(* IEC 61131-3 sources: s7-to-codesys/tests/POUs/Scenarios/FB_AnalogIn_ScenarioTest, 7 files *)

(* ---- FB_AnalogIn_ScenarioTest.decl.st ---- *)
// AUTO-GENERATED — не редактировать: s7conv gen-tests, сценарии scenarios/FB_AnalogIn.csv
// Правка — в CSV (scenarios/README.md), затем python -m s7conv build-corpus.
// Назначение: тесты поведения сконвертированного FB_AnalogIn по сценариям CSV (сценариев: 6, строк: 47):
//             один метод-тест на сценарий, строки — по порядку с моделируемым временем GVL_S7Clock.
//             Ожидаемые значения — из CSV (эталонные модели по описанию логики блока), не из
//             результата конвертации.
// Автор:      s7conv 0.1.0 (сгенерировано)
// Версия:     не указана
// Документ:   scenarios/README.md, docs/methodology.md, раздел «Проверка поведения»
FUNCTION_BLOCK FB_AnalogIn_ScenarioTest EXTENDS coUnit.FB_TestSuite
VAR
    fbScalingPoints : FB_AnalogIn;  // свой экземпляр на сценарий
    xScalingPointsDone : BOOL;  // сценарий выполнен (выполняется один раз)
    fbHighLimitsHysteresis : FB_AnalogIn;  // свой экземпляр на сценарий
    xHighLimitsHysteresisDone : BOOL;  // сценарий выполнен (выполняется один раз)
    fbLowLimitsHysteresis : FB_AnalogIn;  // свой экземпляр на сценарий
    xLowLimitsHysteresisDone : BOOL;  // сценарий выполнен (выполняется один раз)
    fbChannelDiagnostics : FB_AnalogIn;  // свой экземпляр на сценарий
    xChannelDiagnosticsDone : BOOL;  // сценарий выполнен (выполняется один раз)
    fbSimulation : FB_AnalogIn;  // свой экземпляр на сценарий
    xSimulationDone : BOOL;  // сценарий выполнен (выполняется один раз)
    fbCustomRanges : FB_AnalogIn;  // свой экземпляр на сценарий
    xCustomRangesDone : BOOL;  // сценарий выполнен (выполняется один раз)
END_VAR

(* ---- ChannelDiagnostics.method.impl.st ---- *)
// AUTO-GENERATED — не редактировать: scenarios/FB_AnalogIn.csv, сценарий ChannelDiagnostics
coUnit.TEST('ChannelDiagnostics');
IF NOT xChannelDiagnosticsDone THEN
    xChannelDiagnosticsDone := TRUE;
    GVL_S7Clock.xSimulation := TRUE;

    // #1, t = 0 мс — норма 8.0; замещающее значение 5.0
    GVL_S7Clock.tSimNow := T#0MS;
    fbChannelDiagnostics.raw := 13824;
    fbChannelDiagnostics.rangeLow := 0.0;
    fbChannelDiagnostics.rangeHigh := 16.0;
    fbChannelDiagnostics.limitHH := 14.0;
    fbChannelDiagnostics.limitH := 12.0;
    fbChannelDiagnostics.limitL := 2.0;
    fbChannelDiagnostics.limitLL := 1.0;
    fbChannelDiagnostics.hysteresis := 0.5;
    fbChannelDiagnostics.substitute := 5.0;
    fbChannelDiagnostics.simulation := FALSE;
    fbChannelDiagnostics.simValue := 0.0;
    fbChannelDiagnostics();
    AssertEquals_REAL(Expected := 8.0,
                      Actual := fbChannelDiagnostics.value,
                      Delta := 0.001,
                      Message := 'ChannelDiagnostics#1 value');
    AssertEquals_BOOL(Expected := TRUE, Actual := fbChannelDiagnostics.valid, Message := 'ChannelDiagnostics#1 valid');
    AssertEquals_BOOL(Expected := FALSE,
                      Actual := fbChannelDiagnostics.channelFault,
                      Message := 'ChannelDiagnostics#1 channelFault');
    AssertEquals_BOOL(Expected := FALSE,
                      Actual := fbChannelDiagnostics.overrange,
                      Message := 'ChannelDiagnostics#1 overrange');
    AssertEquals_BOOL(Expected := FALSE,
                      Actual := fbChannelDiagnostics.underrange,
                      Message := 'ChannelDiagnostics#1 underrange');
    AssertEquals_BOOL(Expected := FALSE,
                      Actual := fbChannelDiagnostics.alarmHH,
                      Message := 'ChannelDiagnostics#1 alarmHH');
    AssertEquals_BOOL(Expected := FALSE, Actual := fbChannelDiagnostics.warnH, Message := 'ChannelDiagnostics#1 warnH');
    AssertEquals_BOOL(Expected := FALSE, Actual := fbChannelDiagnostics.warnL, Message := 'ChannelDiagnostics#1 warnL');
    AssertEquals_BOOL(Expected := FALSE,
                      Actual := fbChannelDiagnostics.alarmLL,
                      Message := 'ChannelDiagnostics#1 alarmLL');
    AssertEquals_WORD(Expected := 16#0001,
                      Actual := fbChannelDiagnostics.statusWord,
                      Message := 'ChannelDiagnostics#1 statusWord');

    // #2, t = 100 мс — выше номинала: overrange, value ограничено 16.0, HH и H
    GVL_S7Clock.tSimNow := T#100MS;
    fbChannelDiagnostics.raw := 27649;
    fbChannelDiagnostics();
    AssertEquals_REAL(Expected := 16.0,
                      Actual := fbChannelDiagnostics.value,
                      Delta := 0.001,
                      Message := 'ChannelDiagnostics#2 value');
    AssertEquals_BOOL(Expected := TRUE, Actual := fbChannelDiagnostics.valid, Message := 'ChannelDiagnostics#2 valid');
    AssertEquals_BOOL(Expected := FALSE,
                      Actual := fbChannelDiagnostics.channelFault,
                      Message := 'ChannelDiagnostics#2 channelFault');
    AssertEquals_BOOL(Expected := TRUE,
                      Actual := fbChannelDiagnostics.overrange,
                      Message := 'ChannelDiagnostics#2 overrange');
    AssertEquals_BOOL(Expected := FALSE,
                      Actual := fbChannelDiagnostics.underrange,
                      Message := 'ChannelDiagnostics#2 underrange');
    AssertEquals_BOOL(Expected := TRUE,
                      Actual := fbChannelDiagnostics.alarmHH,
                      Message := 'ChannelDiagnostics#2 alarmHH');
    AssertEquals_BOOL(Expected := TRUE, Actual := fbChannelDiagnostics.warnH, Message := 'ChannelDiagnostics#2 warnH');
    AssertEquals_BOOL(Expected := FALSE, Actual := fbChannelDiagnostics.warnL, Message := 'ChannelDiagnostics#2 warnL');
    AssertEquals_BOOL(Expected := FALSE,
                      Actual := fbChannelDiagnostics.alarmLL,
                      Message := 'ChannelDiagnostics#2 alarmLL');
    AssertEquals_WORD(Expected := 16#0035,
                      Actual := fbChannelDiagnostics.statusWord,
                      Message := 'ChannelDiagnostics#2 statusWord');

    // #3, t = 200 мс — верхняя граница зоны перегрузки — ещё не неисправность
    GVL_S7Clock.tSimNow := T#200MS;
    fbChannelDiagnostics.raw := 32511;
    fbChannelDiagnostics();
    AssertEquals_REAL(Expected := 16.0,
                      Actual := fbChannelDiagnostics.value,
                      Delta := 0.001,
                      Message := 'ChannelDiagnostics#3 value');
    AssertEquals_BOOL(Expected := TRUE, Actual := fbChannelDiagnostics.valid, Message := 'ChannelDiagnostics#3 valid');
    AssertEquals_BOOL(Expected := FALSE,
                      Actual := fbChannelDiagnostics.channelFault,
                      Message := 'ChannelDiagnostics#3 channelFault');
    AssertEquals_BOOL(Expected := TRUE,
                      Actual := fbChannelDiagnostics.overrange,
                      Message := 'ChannelDiagnostics#3 overrange');
    AssertEquals_BOOL(Expected := FALSE,
                      Actual := fbChannelDiagnostics.underrange,
                      Message := 'ChannelDiagnostics#3 underrange');
    AssertEquals_BOOL(Expected := TRUE,
                      Actual := fbChannelDiagnostics.alarmHH,
                      Message := 'ChannelDiagnostics#3 alarmHH');
    AssertEquals_BOOL(Expected := TRUE, Actual := fbChannelDiagnostics.warnH, Message := 'ChannelDiagnostics#3 warnH');
    AssertEquals_BOOL(Expected := FALSE, Actual := fbChannelDiagnostics.warnL, Message := 'ChannelDiagnostics#3 warnL');
    AssertEquals_BOOL(Expected := FALSE,
                      Actual := fbChannelDiagnostics.alarmLL,
                      Message := 'ChannelDiagnostics#3 alarmLL');
    AssertEquals_WORD(Expected := 16#0035,
                      Actual := fbChannelDiagnostics.statusWord,
                      Message := 'ChannelDiagnostics#3 statusWord');

    // #4, t = 300 мс — за зоной перегрузки: channelFault, value := substitute, уставки сброшены
    GVL_S7Clock.tSimNow := T#300MS;
    fbChannelDiagnostics.raw := 32512;
    fbChannelDiagnostics();
    AssertEquals_REAL(Expected := 5.0,
                      Actual := fbChannelDiagnostics.value,
                      Delta := 0.001,
                      Message := 'ChannelDiagnostics#4 value');
    AssertEquals_BOOL(Expected := FALSE, Actual := fbChannelDiagnostics.valid, Message := 'ChannelDiagnostics#4 valid');
    AssertEquals_BOOL(Expected := TRUE,
                      Actual := fbChannelDiagnostics.channelFault,
                      Message := 'ChannelDiagnostics#4 channelFault');
    AssertEquals_BOOL(Expected := FALSE,
                      Actual := fbChannelDiagnostics.overrange,
                      Message := 'ChannelDiagnostics#4 overrange');
    AssertEquals_BOOL(Expected := FALSE,
                      Actual := fbChannelDiagnostics.underrange,
                      Message := 'ChannelDiagnostics#4 underrange');
    AssertEquals_BOOL(Expected := FALSE,
                      Actual := fbChannelDiagnostics.alarmHH,
                      Message := 'ChannelDiagnostics#4 alarmHH');
    AssertEquals_BOOL(Expected := FALSE, Actual := fbChannelDiagnostics.warnH, Message := 'ChannelDiagnostics#4 warnH');
    AssertEquals_BOOL(Expected := FALSE, Actual := fbChannelDiagnostics.warnL, Message := 'ChannelDiagnostics#4 warnL');
    AssertEquals_BOOL(Expected := FALSE,
                      Actual := fbChannelDiagnostics.alarmLL,
                      Message := 'ChannelDiagnostics#4 alarmLL');
    AssertEquals_WORD(Expected := 16#0002,
                      Actual := fbChannelDiagnostics.statusWord,
                      Message := 'ChannelDiagnostics#4 statusWord');

    // #5, t = 400 мс — переполнение/обрыв (7FFF)
    GVL_S7Clock.tSimNow := T#400MS;
    fbChannelDiagnostics.raw := 32767;
    fbChannelDiagnostics();
    AssertEquals_REAL(Expected := 5.0,
                      Actual := fbChannelDiagnostics.value,
                      Delta := 0.001,
                      Message := 'ChannelDiagnostics#5 value');
    AssertEquals_BOOL(Expected := FALSE, Actual := fbChannelDiagnostics.valid, Message := 'ChannelDiagnostics#5 valid');
    AssertEquals_BOOL(Expected := TRUE,
                      Actual := fbChannelDiagnostics.channelFault,
                      Message := 'ChannelDiagnostics#5 channelFault');
    AssertEquals_BOOL(Expected := FALSE,
                      Actual := fbChannelDiagnostics.overrange,
                      Message := 'ChannelDiagnostics#5 overrange');
    AssertEquals_BOOL(Expected := FALSE,
                      Actual := fbChannelDiagnostics.underrange,
                      Message := 'ChannelDiagnostics#5 underrange');
    AssertEquals_BOOL(Expected := FALSE,
                      Actual := fbChannelDiagnostics.alarmHH,
                      Message := 'ChannelDiagnostics#5 alarmHH');
    AssertEquals_BOOL(Expected := FALSE, Actual := fbChannelDiagnostics.warnH, Message := 'ChannelDiagnostics#5 warnH');
    AssertEquals_BOOL(Expected := FALSE, Actual := fbChannelDiagnostics.warnL, Message := 'ChannelDiagnostics#5 warnL');
    AssertEquals_BOOL(Expected := FALSE,
                      Actual := fbChannelDiagnostics.alarmLL,
                      Message := 'ChannelDiagnostics#5 alarmLL');
    AssertEquals_WORD(Expected := 16#0002,
                      Actual := fbChannelDiagnostics.statusWord,
                      Message := 'ChannelDiagnostics#5 statusWord');

    // #6, t = 500 мс — канал восстановлен: 8.0, уставки снова считаются (HH не держится)
    GVL_S7Clock.tSimNow := T#500MS;
    fbChannelDiagnostics.raw := 13824;
    fbChannelDiagnostics();
    AssertEquals_REAL(Expected := 8.0,
                      Actual := fbChannelDiagnostics.value,
                      Delta := 0.001,
                      Message := 'ChannelDiagnostics#6 value');
    AssertEquals_BOOL(Expected := TRUE, Actual := fbChannelDiagnostics.valid, Message := 'ChannelDiagnostics#6 valid');
    AssertEquals_BOOL(Expected := FALSE,
                      Actual := fbChannelDiagnostics.channelFault,
                      Message := 'ChannelDiagnostics#6 channelFault');
    AssertEquals_BOOL(Expected := FALSE,
                      Actual := fbChannelDiagnostics.overrange,
                      Message := 'ChannelDiagnostics#6 overrange');
    AssertEquals_BOOL(Expected := FALSE,
                      Actual := fbChannelDiagnostics.underrange,
                      Message := 'ChannelDiagnostics#6 underrange');
    AssertEquals_BOOL(Expected := FALSE,
                      Actual := fbChannelDiagnostics.alarmHH,
                      Message := 'ChannelDiagnostics#6 alarmHH');
    AssertEquals_BOOL(Expected := FALSE, Actual := fbChannelDiagnostics.warnH, Message := 'ChannelDiagnostics#6 warnH');
    AssertEquals_BOOL(Expected := FALSE, Actual := fbChannelDiagnostics.warnL, Message := 'ChannelDiagnostics#6 warnL');
    AssertEquals_BOOL(Expected := FALSE,
                      Actual := fbChannelDiagnostics.alarmLL,
                      Message := 'ChannelDiagnostics#6 alarmLL');
    AssertEquals_WORD(Expected := 16#0001,
                      Actual := fbChannelDiagnostics.statusWord,
                      Message := 'ChannelDiagnostics#6 statusWord');

    // #7, t = 600 мс — ниже номинала: underrange, value ограничено 0.0, L и LL
    GVL_S7Clock.tSimNow := T#600MS;
    fbChannelDiagnostics.raw := -1;
    fbChannelDiagnostics();
    AssertEquals_REAL(Expected := 0.0,
                      Actual := fbChannelDiagnostics.value,
                      Delta := 0.001,
                      Message := 'ChannelDiagnostics#7 value');
    AssertEquals_BOOL(Expected := TRUE, Actual := fbChannelDiagnostics.valid, Message := 'ChannelDiagnostics#7 valid');
    AssertEquals_BOOL(Expected := FALSE,
                      Actual := fbChannelDiagnostics.channelFault,
                      Message := 'ChannelDiagnostics#7 channelFault');
    AssertEquals_BOOL(Expected := FALSE,
                      Actual := fbChannelDiagnostics.overrange,
                      Message := 'ChannelDiagnostics#7 overrange');
    AssertEquals_BOOL(Expected := TRUE,
                      Actual := fbChannelDiagnostics.underrange,
                      Message := 'ChannelDiagnostics#7 underrange');
    AssertEquals_BOOL(Expected := FALSE,
                      Actual := fbChannelDiagnostics.alarmHH,
                      Message := 'ChannelDiagnostics#7 alarmHH');
    AssertEquals_BOOL(Expected := FALSE, Actual := fbChannelDiagnostics.warnH, Message := 'ChannelDiagnostics#7 warnH');
    AssertEquals_BOOL(Expected := TRUE, Actual := fbChannelDiagnostics.warnL, Message := 'ChannelDiagnostics#7 warnL');
    AssertEquals_BOOL(Expected := TRUE,
                      Actual := fbChannelDiagnostics.alarmLL,
                      Message := 'ChannelDiagnostics#7 alarmLL');
    AssertEquals_WORD(Expected := 16#00C9,
                      Actual := fbChannelDiagnostics.statusWord,
                      Message := 'ChannelDiagnostics#7 statusWord');

    // #8, t = 700 мс — нижняя граница зоны перегрузки — ещё не неисправность
    GVL_S7Clock.tSimNow := T#700MS;
    fbChannelDiagnostics.raw := -4864;
    fbChannelDiagnostics();
    AssertEquals_REAL(Expected := 0.0,
                      Actual := fbChannelDiagnostics.value,
                      Delta := 0.001,
                      Message := 'ChannelDiagnostics#8 value');
    AssertEquals_BOOL(Expected := TRUE, Actual := fbChannelDiagnostics.valid, Message := 'ChannelDiagnostics#8 valid');
    AssertEquals_BOOL(Expected := FALSE,
                      Actual := fbChannelDiagnostics.channelFault,
                      Message := 'ChannelDiagnostics#8 channelFault');
    AssertEquals_BOOL(Expected := FALSE,
                      Actual := fbChannelDiagnostics.overrange,
                      Message := 'ChannelDiagnostics#8 overrange');
    AssertEquals_BOOL(Expected := TRUE,
                      Actual := fbChannelDiagnostics.underrange,
                      Message := 'ChannelDiagnostics#8 underrange');
    AssertEquals_BOOL(Expected := FALSE,
                      Actual := fbChannelDiagnostics.alarmHH,
                      Message := 'ChannelDiagnostics#8 alarmHH');
    AssertEquals_BOOL(Expected := FALSE, Actual := fbChannelDiagnostics.warnH, Message := 'ChannelDiagnostics#8 warnH');
    AssertEquals_BOOL(Expected := TRUE, Actual := fbChannelDiagnostics.warnL, Message := 'ChannelDiagnostics#8 warnL');
    AssertEquals_BOOL(Expected := TRUE,
                      Actual := fbChannelDiagnostics.alarmLL,
                      Message := 'ChannelDiagnostics#8 alarmLL');
    AssertEquals_WORD(Expected := 16#00C9,
                      Actual := fbChannelDiagnostics.statusWord,
                      Message := 'ChannelDiagnostics#8 statusWord');

    // #9, t = 800 мс — за зоной: channelFault
    GVL_S7Clock.tSimNow := T#800MS;
    fbChannelDiagnostics.raw := -4865;
    fbChannelDiagnostics();
    AssertEquals_REAL(Expected := 5.0,
                      Actual := fbChannelDiagnostics.value,
                      Delta := 0.001,
                      Message := 'ChannelDiagnostics#9 value');
    AssertEquals_BOOL(Expected := FALSE, Actual := fbChannelDiagnostics.valid, Message := 'ChannelDiagnostics#9 valid');
    AssertEquals_BOOL(Expected := TRUE,
                      Actual := fbChannelDiagnostics.channelFault,
                      Message := 'ChannelDiagnostics#9 channelFault');
    AssertEquals_BOOL(Expected := FALSE,
                      Actual := fbChannelDiagnostics.overrange,
                      Message := 'ChannelDiagnostics#9 overrange');
    AssertEquals_BOOL(Expected := FALSE,
                      Actual := fbChannelDiagnostics.underrange,
                      Message := 'ChannelDiagnostics#9 underrange');
    AssertEquals_BOOL(Expected := FALSE,
                      Actual := fbChannelDiagnostics.alarmHH,
                      Message := 'ChannelDiagnostics#9 alarmHH');
    AssertEquals_BOOL(Expected := FALSE, Actual := fbChannelDiagnostics.warnH, Message := 'ChannelDiagnostics#9 warnH');
    AssertEquals_BOOL(Expected := FALSE, Actual := fbChannelDiagnostics.warnL, Message := 'ChannelDiagnostics#9 warnL');
    AssertEquals_BOOL(Expected := FALSE,
                      Actual := fbChannelDiagnostics.alarmLL,
                      Message := 'ChannelDiagnostics#9 alarmLL');
    AssertEquals_WORD(Expected := 16#0002,
                      Actual := fbChannelDiagnostics.statusWord,
                      Message := 'ChannelDiagnostics#9 statusWord');

    // #10, t = 900 мс — антипереполнение (8000)
    GVL_S7Clock.tSimNow := T#900MS;
    fbChannelDiagnostics.raw := -32768;
    fbChannelDiagnostics();
    AssertEquals_REAL(Expected := 5.0,
                      Actual := fbChannelDiagnostics.value,
                      Delta := 0.001,
                      Message := 'ChannelDiagnostics#10 value');
    AssertEquals_BOOL(Expected := FALSE,
                      Actual := fbChannelDiagnostics.valid,
                      Message := 'ChannelDiagnostics#10 valid');
    AssertEquals_BOOL(Expected := TRUE,
                      Actual := fbChannelDiagnostics.channelFault,
                      Message := 'ChannelDiagnostics#10 channelFault');
    AssertEquals_BOOL(Expected := FALSE,
                      Actual := fbChannelDiagnostics.overrange,
                      Message := 'ChannelDiagnostics#10 overrange');
    AssertEquals_BOOL(Expected := FALSE,
                      Actual := fbChannelDiagnostics.underrange,
                      Message := 'ChannelDiagnostics#10 underrange');
    AssertEquals_BOOL(Expected := FALSE,
                      Actual := fbChannelDiagnostics.alarmHH,
                      Message := 'ChannelDiagnostics#10 alarmHH');
    AssertEquals_BOOL(Expected := FALSE,
                      Actual := fbChannelDiagnostics.warnH,
                      Message := 'ChannelDiagnostics#10 warnH');
    AssertEquals_BOOL(Expected := FALSE,
                      Actual := fbChannelDiagnostics.warnL,
                      Message := 'ChannelDiagnostics#10 warnL');
    AssertEquals_BOOL(Expected := FALSE,
                      Actual := fbChannelDiagnostics.alarmLL,
                      Message := 'ChannelDiagnostics#10 alarmLL');
    AssertEquals_WORD(Expected := 16#0002,
                      Actual := fbChannelDiagnostics.statusWord,
                      Message := 'ChannelDiagnostics#10 statusWord');

    // #11, t = 1000 мс — канал восстановлен: 2.0 — только L
    GVL_S7Clock.tSimNow := T#1000MS;
    fbChannelDiagnostics.raw := 3456;
    fbChannelDiagnostics();
    AssertEquals_REAL(Expected := 2.0,
                      Actual := fbChannelDiagnostics.value,
                      Delta := 0.001,
                      Message := 'ChannelDiagnostics#11 value');
    AssertEquals_BOOL(Expected := TRUE, Actual := fbChannelDiagnostics.valid, Message := 'ChannelDiagnostics#11 valid');
    AssertEquals_BOOL(Expected := FALSE,
                      Actual := fbChannelDiagnostics.channelFault,
                      Message := 'ChannelDiagnostics#11 channelFault');
    AssertEquals_BOOL(Expected := FALSE,
                      Actual := fbChannelDiagnostics.overrange,
                      Message := 'ChannelDiagnostics#11 overrange');
    AssertEquals_BOOL(Expected := FALSE,
                      Actual := fbChannelDiagnostics.underrange,
                      Message := 'ChannelDiagnostics#11 underrange');
    AssertEquals_BOOL(Expected := FALSE,
                      Actual := fbChannelDiagnostics.alarmHH,
                      Message := 'ChannelDiagnostics#11 alarmHH');
    AssertEquals_BOOL(Expected := FALSE,
                      Actual := fbChannelDiagnostics.warnH,
                      Message := 'ChannelDiagnostics#11 warnH');
    AssertEquals_BOOL(Expected := TRUE, Actual := fbChannelDiagnostics.warnL, Message := 'ChannelDiagnostics#11 warnL');
    AssertEquals_BOOL(Expected := FALSE,
                      Actual := fbChannelDiagnostics.alarmLL,
                      Message := 'ChannelDiagnostics#11 alarmLL');
    AssertEquals_WORD(Expected := 16#0041,
                      Actual := fbChannelDiagnostics.statusWord,
                      Message := 'ChannelDiagnostics#11 statusWord');

    GVL_S7Clock.xSimulation := FALSE;
END_IF
coUnit.TEST_FINISHED();

(* ---- CustomRanges.method.impl.st ---- *)
// AUTO-GENERATED — не редактировать: scenarios/FB_AnalogIn.csv, сценарий CustomRanges
coUnit.TEST('CustomRanges');
IF NOT xCustomRangesDone THEN
    xCustomRangesDone := TRUE;
    GVL_S7Clock.xSimulation := TRUE;

    // #1, t = 0 мс — шкала -50...150: четверть -> 0.0 = limitL
    GVL_S7Clock.tSimNow := T#0MS;
    fbCustomRanges.raw := 6912;
    fbCustomRanges.rangeLow := -50.0;
    fbCustomRanges.rangeHigh := 150.0;
    fbCustomRanges.limitHH := 120.0;
    fbCustomRanges.limitH := 100.0;
    fbCustomRanges.limitL := 0.0;
    fbCustomRanges.limitLL := -20.0;
    fbCustomRanges.hysteresis := 2.0;
    fbCustomRanges.substitute := 0.0;
    fbCustomRanges.simulation := FALSE;
    fbCustomRanges.simValue := 0.0;
    fbCustomRanges();
    AssertEquals_REAL(Expected := 0.0,
                      Actual := fbCustomRanges.value,
                      Delta := 0.001,
                      Message := 'CustomRanges#1 value');
    AssertEquals_BOOL(Expected := TRUE, Actual := fbCustomRanges.valid, Message := 'CustomRanges#1 valid');
    AssertEquals_BOOL(Expected := FALSE,
                      Actual := fbCustomRanges.channelFault,
                      Message := 'CustomRanges#1 channelFault');
    AssertEquals_BOOL(Expected := FALSE, Actual := fbCustomRanges.overrange, Message := 'CustomRanges#1 overrange');
    AssertEquals_BOOL(Expected := FALSE, Actual := fbCustomRanges.underrange, Message := 'CustomRanges#1 underrange');
    AssertEquals_BOOL(Expected := FALSE, Actual := fbCustomRanges.alarmHH, Message := 'CustomRanges#1 alarmHH');
    AssertEquals_BOOL(Expected := FALSE, Actual := fbCustomRanges.warnH, Message := 'CustomRanges#1 warnH');
    AssertEquals_BOOL(Expected := TRUE, Actual := fbCustomRanges.warnL, Message := 'CustomRanges#1 warnL');
    AssertEquals_BOOL(Expected := FALSE, Actual := fbCustomRanges.alarmLL, Message := 'CustomRanges#1 alarmLL');
    AssertEquals_WORD(Expected := 16#0041, Actual := fbCustomRanges.statusWord, Message := 'CustomRanges#1 statusWord');

    // #2, t = 100 мс — три четверти -> 100.0 = limitH; L сброшен
    GVL_S7Clock.tSimNow := T#100MS;
    fbCustomRanges.raw := 20736;
    fbCustomRanges();
    AssertEquals_REAL(Expected := 100.0,
                      Actual := fbCustomRanges.value,
                      Delta := 0.001,
                      Message := 'CustomRanges#2 value');
    AssertEquals_BOOL(Expected := TRUE, Actual := fbCustomRanges.valid, Message := 'CustomRanges#2 valid');
    AssertEquals_BOOL(Expected := FALSE,
                      Actual := fbCustomRanges.channelFault,
                      Message := 'CustomRanges#2 channelFault');
    AssertEquals_BOOL(Expected := FALSE, Actual := fbCustomRanges.overrange, Message := 'CustomRanges#2 overrange');
    AssertEquals_BOOL(Expected := FALSE, Actual := fbCustomRanges.underrange, Message := 'CustomRanges#2 underrange');
    AssertEquals_BOOL(Expected := FALSE, Actual := fbCustomRanges.alarmHH, Message := 'CustomRanges#2 alarmHH');
    AssertEquals_BOOL(Expected := TRUE, Actual := fbCustomRanges.warnH, Message := 'CustomRanges#2 warnH');
    AssertEquals_BOOL(Expected := FALSE, Actual := fbCustomRanges.warnL, Message := 'CustomRanges#2 warnL');
    AssertEquals_BOOL(Expected := FALSE, Actual := fbCustomRanges.alarmLL, Message := 'CustomRanges#2 alarmLL');
    AssertEquals_WORD(Expected := 16#0021, Actual := fbCustomRanges.statusWord, Message := 'CustomRanges#2 statusWord');

    // #3, t = 200 мс — максимум -> 150.0: HH и H
    GVL_S7Clock.tSimNow := T#200MS;
    fbCustomRanges.raw := 27648;
    fbCustomRanges();
    AssertEquals_REAL(Expected := 150.0,
                      Actual := fbCustomRanges.value,
                      Delta := 0.001,
                      Message := 'CustomRanges#3 value');
    AssertEquals_BOOL(Expected := TRUE, Actual := fbCustomRanges.valid, Message := 'CustomRanges#3 valid');
    AssertEquals_BOOL(Expected := FALSE,
                      Actual := fbCustomRanges.channelFault,
                      Message := 'CustomRanges#3 channelFault');
    AssertEquals_BOOL(Expected := FALSE, Actual := fbCustomRanges.overrange, Message := 'CustomRanges#3 overrange');
    AssertEquals_BOOL(Expected := FALSE, Actual := fbCustomRanges.underrange, Message := 'CustomRanges#3 underrange');
    AssertEquals_BOOL(Expected := TRUE, Actual := fbCustomRanges.alarmHH, Message := 'CustomRanges#3 alarmHH');
    AssertEquals_BOOL(Expected := TRUE, Actual := fbCustomRanges.warnH, Message := 'CustomRanges#3 warnH');
    AssertEquals_BOOL(Expected := FALSE, Actual := fbCustomRanges.warnL, Message := 'CustomRanges#3 warnL');
    AssertEquals_BOOL(Expected := FALSE, Actual := fbCustomRanges.alarmLL, Message := 'CustomRanges#3 alarmLL');
    AssertEquals_WORD(Expected := 16#0031, Actual := fbCustomRanges.statusWord, Message := 'CustomRanges#3 statusWord');

    // #4, t = 300 мс — минимум -> -50.0: L и LL
    GVL_S7Clock.tSimNow := T#300MS;
    fbCustomRanges.raw := 0;
    fbCustomRanges();
    AssertEquals_REAL(Expected := -50.0,
                      Actual := fbCustomRanges.value,
                      Delta := 0.001,
                      Message := 'CustomRanges#4 value');
    AssertEquals_BOOL(Expected := TRUE, Actual := fbCustomRanges.valid, Message := 'CustomRanges#4 valid');
    AssertEquals_BOOL(Expected := FALSE,
                      Actual := fbCustomRanges.channelFault,
                      Message := 'CustomRanges#4 channelFault');
    AssertEquals_BOOL(Expected := FALSE, Actual := fbCustomRanges.overrange, Message := 'CustomRanges#4 overrange');
    AssertEquals_BOOL(Expected := FALSE, Actual := fbCustomRanges.underrange, Message := 'CustomRanges#4 underrange');
    AssertEquals_BOOL(Expected := FALSE, Actual := fbCustomRanges.alarmHH, Message := 'CustomRanges#4 alarmHH');
    AssertEquals_BOOL(Expected := FALSE, Actual := fbCustomRanges.warnH, Message := 'CustomRanges#4 warnH');
    AssertEquals_BOOL(Expected := TRUE, Actual := fbCustomRanges.warnL, Message := 'CustomRanges#4 warnL');
    AssertEquals_BOOL(Expected := TRUE, Actual := fbCustomRanges.alarmLL, Message := 'CustomRanges#4 alarmLL');
    AssertEquals_WORD(Expected := 16#00C1, Actual := fbCustomRanges.statusWord, Message := 'CustomRanges#4 statusWord');

    // #5, t = 400 мс — обратная шкала 16...0: четверть -> 12.0 = limitH
    GVL_S7Clock.tSimNow := T#400MS;
    fbCustomRanges.raw := 6912;
    fbCustomRanges.rangeLow := 16.0;
    fbCustomRanges.rangeHigh := 0.0;
    fbCustomRanges.limitHH := 14.0;
    fbCustomRanges.limitH := 12.0;
    fbCustomRanges.limitL := 2.0;
    fbCustomRanges.limitLL := 1.0;
    fbCustomRanges.hysteresis := 0.5;
    fbCustomRanges();
    AssertEquals_REAL(Expected := 12.0,
                      Actual := fbCustomRanges.value,
                      Delta := 0.001,
                      Message := 'CustomRanges#5 value');
    AssertEquals_BOOL(Expected := TRUE, Actual := fbCustomRanges.valid, Message := 'CustomRanges#5 valid');
    AssertEquals_BOOL(Expected := FALSE,
                      Actual := fbCustomRanges.channelFault,
                      Message := 'CustomRanges#5 channelFault');
    AssertEquals_BOOL(Expected := FALSE, Actual := fbCustomRanges.overrange, Message := 'CustomRanges#5 overrange');
    AssertEquals_BOOL(Expected := FALSE, Actual := fbCustomRanges.underrange, Message := 'CustomRanges#5 underrange');
    AssertEquals_BOOL(Expected := FALSE, Actual := fbCustomRanges.alarmHH, Message := 'CustomRanges#5 alarmHH');
    AssertEquals_BOOL(Expected := TRUE, Actual := fbCustomRanges.warnH, Message := 'CustomRanges#5 warnH');
    AssertEquals_BOOL(Expected := FALSE, Actual := fbCustomRanges.warnL, Message := 'CustomRanges#5 warnL');
    AssertEquals_BOOL(Expected := FALSE, Actual := fbCustomRanges.alarmLL, Message := 'CustomRanges#5 alarmLL');
    AssertEquals_WORD(Expected := 16#0021, Actual := fbCustomRanges.statusWord, Message := 'CustomRanges#5 statusWord');

    // #6, t = 500 мс — обратная шкала: максимум raw -> 0.0, L и LL
    GVL_S7Clock.tSimNow := T#500MS;
    fbCustomRanges.raw := 27648;
    fbCustomRanges();
    AssertEquals_REAL(Expected := 0.0,
                      Actual := fbCustomRanges.value,
                      Delta := 0.001,
                      Message := 'CustomRanges#6 value');
    AssertEquals_BOOL(Expected := TRUE, Actual := fbCustomRanges.valid, Message := 'CustomRanges#6 valid');
    AssertEquals_BOOL(Expected := FALSE,
                      Actual := fbCustomRanges.channelFault,
                      Message := 'CustomRanges#6 channelFault');
    AssertEquals_BOOL(Expected := FALSE, Actual := fbCustomRanges.overrange, Message := 'CustomRanges#6 overrange');
    AssertEquals_BOOL(Expected := FALSE, Actual := fbCustomRanges.underrange, Message := 'CustomRanges#6 underrange');
    AssertEquals_BOOL(Expected := FALSE, Actual := fbCustomRanges.alarmHH, Message := 'CustomRanges#6 alarmHH');
    AssertEquals_BOOL(Expected := FALSE, Actual := fbCustomRanges.warnH, Message := 'CustomRanges#6 warnH');
    AssertEquals_BOOL(Expected := TRUE, Actual := fbCustomRanges.warnL, Message := 'CustomRanges#6 warnL');
    AssertEquals_BOOL(Expected := TRUE, Actual := fbCustomRanges.alarmLL, Message := 'CustomRanges#6 alarmLL');
    AssertEquals_WORD(Expected := 16#00C1, Actual := fbCustomRanges.statusWord, Message := 'CustomRanges#6 statusWord');

    GVL_S7Clock.xSimulation := FALSE;
END_IF
coUnit.TEST_FINISHED();

(* ---- HighLimitsHysteresis.method.impl.st ---- *)
// AUTO-GENERATED — не редактировать: scenarios/FB_AnalogIn.csv, сценарий HighLimitsHysteresis
coUnit.TEST('HighLimitsHysteresis');
IF NOT xHighLimitsHysteresisDone THEN
    xHighLimitsHysteresisDone := TRUE;
    GVL_S7Clock.xSimulation := TRUE;

    // #1, t = 0 мс — 11.0 — ниже всех верхних уставок
    GVL_S7Clock.tSimNow := T#0MS;
    fbHighLimitsHysteresis.raw := 19008;
    fbHighLimitsHysteresis.rangeLow := 0.0;
    fbHighLimitsHysteresis.rangeHigh := 16.0;
    fbHighLimitsHysteresis.limitHH := 14.0;
    fbHighLimitsHysteresis.limitH := 12.0;
    fbHighLimitsHysteresis.limitL := 2.0;
    fbHighLimitsHysteresis.limitLL := 1.0;
    fbHighLimitsHysteresis.hysteresis := 0.5;
    fbHighLimitsHysteresis.substitute := 0.0;
    fbHighLimitsHysteresis.simulation := FALSE;
    fbHighLimitsHysteresis.simValue := 0.0;
    fbHighLimitsHysteresis();
    AssertEquals_REAL(Expected := 11.0,
                      Actual := fbHighLimitsHysteresis.value,
                      Delta := 0.001,
                      Message := 'HighLimitsHysteresis#1 value');
    AssertEquals_BOOL(Expected := TRUE,
                      Actual := fbHighLimitsHysteresis.valid,
                      Message := 'HighLimitsHysteresis#1 valid');
    AssertEquals_BOOL(Expected := FALSE,
                      Actual := fbHighLimitsHysteresis.channelFault,
                      Message := 'HighLimitsHysteresis#1 channelFault');
    AssertEquals_BOOL(Expected := FALSE,
                      Actual := fbHighLimitsHysteresis.overrange,
                      Message := 'HighLimitsHysteresis#1 overrange');
    AssertEquals_BOOL(Expected := FALSE,
                      Actual := fbHighLimitsHysteresis.underrange,
                      Message := 'HighLimitsHysteresis#1 underrange');
    AssertEquals_BOOL(Expected := FALSE,
                      Actual := fbHighLimitsHysteresis.alarmHH,
                      Message := 'HighLimitsHysteresis#1 alarmHH');
    AssertEquals_BOOL(Expected := FALSE,
                      Actual := fbHighLimitsHysteresis.warnH,
                      Message := 'HighLimitsHysteresis#1 warnH');
    AssertEquals_BOOL(Expected := FALSE,
                      Actual := fbHighLimitsHysteresis.warnL,
                      Message := 'HighLimitsHysteresis#1 warnL');
    AssertEquals_BOOL(Expected := FALSE,
                      Actual := fbHighLimitsHysteresis.alarmLL,
                      Message := 'HighLimitsHysteresis#1 alarmLL');
    AssertEquals_WORD(Expected := 16#0001,
                      Actual := fbHighLimitsHysteresis.statusWord,
                      Message := 'HighLimitsHysteresis#1 statusWord');

    // #2, t = 100 мс — 12.0 = limitH: H включается
    GVL_S7Clock.tSimNow := T#100MS;
    fbHighLimitsHysteresis.raw := 20736;
    fbHighLimitsHysteresis();
    AssertEquals_REAL(Expected := 12.0,
                      Actual := fbHighLimitsHysteresis.value,
                      Delta := 0.001,
                      Message := 'HighLimitsHysteresis#2 value');
    AssertEquals_BOOL(Expected := TRUE,
                      Actual := fbHighLimitsHysteresis.valid,
                      Message := 'HighLimitsHysteresis#2 valid');
    AssertEquals_BOOL(Expected := FALSE,
                      Actual := fbHighLimitsHysteresis.channelFault,
                      Message := 'HighLimitsHysteresis#2 channelFault');
    AssertEquals_BOOL(Expected := FALSE,
                      Actual := fbHighLimitsHysteresis.overrange,
                      Message := 'HighLimitsHysteresis#2 overrange');
    AssertEquals_BOOL(Expected := FALSE,
                      Actual := fbHighLimitsHysteresis.underrange,
                      Message := 'HighLimitsHysteresis#2 underrange');
    AssertEquals_BOOL(Expected := FALSE,
                      Actual := fbHighLimitsHysteresis.alarmHH,
                      Message := 'HighLimitsHysteresis#2 alarmHH');
    AssertEquals_BOOL(Expected := TRUE,
                      Actual := fbHighLimitsHysteresis.warnH,
                      Message := 'HighLimitsHysteresis#2 warnH');
    AssertEquals_BOOL(Expected := FALSE,
                      Actual := fbHighLimitsHysteresis.warnL,
                      Message := 'HighLimitsHysteresis#2 warnL');
    AssertEquals_BOOL(Expected := FALSE,
                      Actual := fbHighLimitsHysteresis.alarmLL,
                      Message := 'HighLimitsHysteresis#2 alarmLL');
    AssertEquals_WORD(Expected := 16#0021,
                      Actual := fbHighLimitsHysteresis.statusWord,
                      Message := 'HighLimitsHysteresis#2 statusWord');

    // #3, t = 200 мс — 11.75 — в зоне гистерезиса, H держится
    GVL_S7Clock.tSimNow := T#200MS;
    fbHighLimitsHysteresis.raw := 20304;
    fbHighLimitsHysteresis();
    AssertEquals_REAL(Expected := 11.75,
                      Actual := fbHighLimitsHysteresis.value,
                      Delta := 0.001,
                      Message := 'HighLimitsHysteresis#3 value');
    AssertEquals_BOOL(Expected := TRUE,
                      Actual := fbHighLimitsHysteresis.valid,
                      Message := 'HighLimitsHysteresis#3 valid');
    AssertEquals_BOOL(Expected := FALSE,
                      Actual := fbHighLimitsHysteresis.channelFault,
                      Message := 'HighLimitsHysteresis#3 channelFault');
    AssertEquals_BOOL(Expected := FALSE,
                      Actual := fbHighLimitsHysteresis.overrange,
                      Message := 'HighLimitsHysteresis#3 overrange');
    AssertEquals_BOOL(Expected := FALSE,
                      Actual := fbHighLimitsHysteresis.underrange,
                      Message := 'HighLimitsHysteresis#3 underrange');
    AssertEquals_BOOL(Expected := FALSE,
                      Actual := fbHighLimitsHysteresis.alarmHH,
                      Message := 'HighLimitsHysteresis#3 alarmHH');
    AssertEquals_BOOL(Expected := TRUE,
                      Actual := fbHighLimitsHysteresis.warnH,
                      Message := 'HighLimitsHysteresis#3 warnH');
    AssertEquals_BOOL(Expected := FALSE,
                      Actual := fbHighLimitsHysteresis.warnL,
                      Message := 'HighLimitsHysteresis#3 warnL');
    AssertEquals_BOOL(Expected := FALSE,
                      Actual := fbHighLimitsHysteresis.alarmLL,
                      Message := 'HighLimitsHysteresis#3 alarmLL');
    AssertEquals_WORD(Expected := 16#0021,
                      Actual := fbHighLimitsHysteresis.statusWord,
                      Message := 'HighLimitsHysteresis#3 statusWord');

    // #4, t = 300 мс — 11.5 = limitH - hysteresis: не меньше порога, H держится
    GVL_S7Clock.tSimNow := T#300MS;
    fbHighLimitsHysteresis.raw := 19872;
    fbHighLimitsHysteresis();
    AssertEquals_REAL(Expected := 11.5,
                      Actual := fbHighLimitsHysteresis.value,
                      Delta := 0.001,
                      Message := 'HighLimitsHysteresis#4 value');
    AssertEquals_BOOL(Expected := TRUE,
                      Actual := fbHighLimitsHysteresis.valid,
                      Message := 'HighLimitsHysteresis#4 valid');
    AssertEquals_BOOL(Expected := FALSE,
                      Actual := fbHighLimitsHysteresis.channelFault,
                      Message := 'HighLimitsHysteresis#4 channelFault');
    AssertEquals_BOOL(Expected := FALSE,
                      Actual := fbHighLimitsHysteresis.overrange,
                      Message := 'HighLimitsHysteresis#4 overrange');
    AssertEquals_BOOL(Expected := FALSE,
                      Actual := fbHighLimitsHysteresis.underrange,
                      Message := 'HighLimitsHysteresis#4 underrange');
    AssertEquals_BOOL(Expected := FALSE,
                      Actual := fbHighLimitsHysteresis.alarmHH,
                      Message := 'HighLimitsHysteresis#4 alarmHH');
    AssertEquals_BOOL(Expected := TRUE,
                      Actual := fbHighLimitsHysteresis.warnH,
                      Message := 'HighLimitsHysteresis#4 warnH');
    AssertEquals_BOOL(Expected := FALSE,
                      Actual := fbHighLimitsHysteresis.warnL,
                      Message := 'HighLimitsHysteresis#4 warnL');
    AssertEquals_BOOL(Expected := FALSE,
                      Actual := fbHighLimitsHysteresis.alarmLL,
                      Message := 'HighLimitsHysteresis#4 alarmLL');
    AssertEquals_WORD(Expected := 16#0021,
                      Actual := fbHighLimitsHysteresis.statusWord,
                      Message := 'HighLimitsHysteresis#4 statusWord');

    // #5, t = 400 мс — 11.25 < 11.5: H сбрасывается
    GVL_S7Clock.tSimNow := T#400MS;
    fbHighLimitsHysteresis.raw := 19440;
    fbHighLimitsHysteresis();
    AssertEquals_REAL(Expected := 11.25,
                      Actual := fbHighLimitsHysteresis.value,
                      Delta := 0.001,
                      Message := 'HighLimitsHysteresis#5 value');
    AssertEquals_BOOL(Expected := TRUE,
                      Actual := fbHighLimitsHysteresis.valid,
                      Message := 'HighLimitsHysteresis#5 valid');
    AssertEquals_BOOL(Expected := FALSE,
                      Actual := fbHighLimitsHysteresis.channelFault,
                      Message := 'HighLimitsHysteresis#5 channelFault');
    AssertEquals_BOOL(Expected := FALSE,
                      Actual := fbHighLimitsHysteresis.overrange,
                      Message := 'HighLimitsHysteresis#5 overrange');
    AssertEquals_BOOL(Expected := FALSE,
                      Actual := fbHighLimitsHysteresis.underrange,
                      Message := 'HighLimitsHysteresis#5 underrange');
    AssertEquals_BOOL(Expected := FALSE,
                      Actual := fbHighLimitsHysteresis.alarmHH,
                      Message := 'HighLimitsHysteresis#5 alarmHH');
    AssertEquals_BOOL(Expected := FALSE,
                      Actual := fbHighLimitsHysteresis.warnH,
                      Message := 'HighLimitsHysteresis#5 warnH');
    AssertEquals_BOOL(Expected := FALSE,
                      Actual := fbHighLimitsHysteresis.warnL,
                      Message := 'HighLimitsHysteresis#5 warnL');
    AssertEquals_BOOL(Expected := FALSE,
                      Actual := fbHighLimitsHysteresis.alarmLL,
                      Message := 'HighLimitsHysteresis#5 alarmLL');
    AssertEquals_WORD(Expected := 16#0001,
                      Actual := fbHighLimitsHysteresis.statusWord,
                      Message := 'HighLimitsHysteresis#5 statusWord');

    // #6, t = 500 мс — 14.0 = limitHH: HH и H
    GVL_S7Clock.tSimNow := T#500MS;
    fbHighLimitsHysteresis.raw := 24192;
    fbHighLimitsHysteresis();
    AssertEquals_REAL(Expected := 14.0,
                      Actual := fbHighLimitsHysteresis.value,
                      Delta := 0.001,
                      Message := 'HighLimitsHysteresis#6 value');
    AssertEquals_BOOL(Expected := TRUE,
                      Actual := fbHighLimitsHysteresis.valid,
                      Message := 'HighLimitsHysteresis#6 valid');
    AssertEquals_BOOL(Expected := FALSE,
                      Actual := fbHighLimitsHysteresis.channelFault,
                      Message := 'HighLimitsHysteresis#6 channelFault');
    AssertEquals_BOOL(Expected := FALSE,
                      Actual := fbHighLimitsHysteresis.overrange,
                      Message := 'HighLimitsHysteresis#6 overrange');
    AssertEquals_BOOL(Expected := FALSE,
                      Actual := fbHighLimitsHysteresis.underrange,
                      Message := 'HighLimitsHysteresis#6 underrange');
    AssertEquals_BOOL(Expected := TRUE,
                      Actual := fbHighLimitsHysteresis.alarmHH,
                      Message := 'HighLimitsHysteresis#6 alarmHH');
    AssertEquals_BOOL(Expected := TRUE,
                      Actual := fbHighLimitsHysteresis.warnH,
                      Message := 'HighLimitsHysteresis#6 warnH');
    AssertEquals_BOOL(Expected := FALSE,
                      Actual := fbHighLimitsHysteresis.warnL,
                      Message := 'HighLimitsHysteresis#6 warnL');
    AssertEquals_BOOL(Expected := FALSE,
                      Actual := fbHighLimitsHysteresis.alarmLL,
                      Message := 'HighLimitsHysteresis#6 alarmLL');
    AssertEquals_WORD(Expected := 16#0031,
                      Actual := fbHighLimitsHysteresis.statusWord,
                      Message := 'HighLimitsHysteresis#6 statusWord');

    // #7, t = 600 мс — 13.5 = limitHH - hysteresis: HH держится
    GVL_S7Clock.tSimNow := T#600MS;
    fbHighLimitsHysteresis.raw := 23328;
    fbHighLimitsHysteresis();
    AssertEquals_REAL(Expected := 13.5,
                      Actual := fbHighLimitsHysteresis.value,
                      Delta := 0.001,
                      Message := 'HighLimitsHysteresis#7 value');
    AssertEquals_BOOL(Expected := TRUE,
                      Actual := fbHighLimitsHysteresis.valid,
                      Message := 'HighLimitsHysteresis#7 valid');
    AssertEquals_BOOL(Expected := FALSE,
                      Actual := fbHighLimitsHysteresis.channelFault,
                      Message := 'HighLimitsHysteresis#7 channelFault');
    AssertEquals_BOOL(Expected := FALSE,
                      Actual := fbHighLimitsHysteresis.overrange,
                      Message := 'HighLimitsHysteresis#7 overrange');
    AssertEquals_BOOL(Expected := FALSE,
                      Actual := fbHighLimitsHysteresis.underrange,
                      Message := 'HighLimitsHysteresis#7 underrange');
    AssertEquals_BOOL(Expected := TRUE,
                      Actual := fbHighLimitsHysteresis.alarmHH,
                      Message := 'HighLimitsHysteresis#7 alarmHH');
    AssertEquals_BOOL(Expected := TRUE,
                      Actual := fbHighLimitsHysteresis.warnH,
                      Message := 'HighLimitsHysteresis#7 warnH');
    AssertEquals_BOOL(Expected := FALSE,
                      Actual := fbHighLimitsHysteresis.warnL,
                      Message := 'HighLimitsHysteresis#7 warnL');
    AssertEquals_BOOL(Expected := FALSE,
                      Actual := fbHighLimitsHysteresis.alarmLL,
                      Message := 'HighLimitsHysteresis#7 alarmLL');
    AssertEquals_WORD(Expected := 16#0031,
                      Actual := fbHighLimitsHysteresis.statusWord,
                      Message := 'HighLimitsHysteresis#7 statusWord');

    // #8, t = 700 мс — 13.25 < 13.5: HH сброшен, H держится
    GVL_S7Clock.tSimNow := T#700MS;
    fbHighLimitsHysteresis.raw := 22896;
    fbHighLimitsHysteresis();
    AssertEquals_REAL(Expected := 13.25,
                      Actual := fbHighLimitsHysteresis.value,
                      Delta := 0.001,
                      Message := 'HighLimitsHysteresis#8 value');
    AssertEquals_BOOL(Expected := TRUE,
                      Actual := fbHighLimitsHysteresis.valid,
                      Message := 'HighLimitsHysteresis#8 valid');
    AssertEquals_BOOL(Expected := FALSE,
                      Actual := fbHighLimitsHysteresis.channelFault,
                      Message := 'HighLimitsHysteresis#8 channelFault');
    AssertEquals_BOOL(Expected := FALSE,
                      Actual := fbHighLimitsHysteresis.overrange,
                      Message := 'HighLimitsHysteresis#8 overrange');
    AssertEquals_BOOL(Expected := FALSE,
                      Actual := fbHighLimitsHysteresis.underrange,
                      Message := 'HighLimitsHysteresis#8 underrange');
    AssertEquals_BOOL(Expected := FALSE,
                      Actual := fbHighLimitsHysteresis.alarmHH,
                      Message := 'HighLimitsHysteresis#8 alarmHH');
    AssertEquals_BOOL(Expected := TRUE,
                      Actual := fbHighLimitsHysteresis.warnH,
                      Message := 'HighLimitsHysteresis#8 warnH');
    AssertEquals_BOOL(Expected := FALSE,
                      Actual := fbHighLimitsHysteresis.warnL,
                      Message := 'HighLimitsHysteresis#8 warnL');
    AssertEquals_BOOL(Expected := FALSE,
                      Actual := fbHighLimitsHysteresis.alarmLL,
                      Message := 'HighLimitsHysteresis#8 alarmLL');
    AssertEquals_WORD(Expected := 16#0021,
                      Actual := fbHighLimitsHysteresis.statusWord,
                      Message := 'HighLimitsHysteresis#8 statusWord');

    // #9, t = 800 мс — 13.75 < 14.0: HH снова не включается
    GVL_S7Clock.tSimNow := T#800MS;
    fbHighLimitsHysteresis.raw := 23760;
    fbHighLimitsHysteresis();
    AssertEquals_REAL(Expected := 13.75,
                      Actual := fbHighLimitsHysteresis.value,
                      Delta := 0.001,
                      Message := 'HighLimitsHysteresis#9 value');
    AssertEquals_BOOL(Expected := TRUE,
                      Actual := fbHighLimitsHysteresis.valid,
                      Message := 'HighLimitsHysteresis#9 valid');
    AssertEquals_BOOL(Expected := FALSE,
                      Actual := fbHighLimitsHysteresis.channelFault,
                      Message := 'HighLimitsHysteresis#9 channelFault');
    AssertEquals_BOOL(Expected := FALSE,
                      Actual := fbHighLimitsHysteresis.overrange,
                      Message := 'HighLimitsHysteresis#9 overrange');
    AssertEquals_BOOL(Expected := FALSE,
                      Actual := fbHighLimitsHysteresis.underrange,
                      Message := 'HighLimitsHysteresis#9 underrange');
    AssertEquals_BOOL(Expected := FALSE,
                      Actual := fbHighLimitsHysteresis.alarmHH,
                      Message := 'HighLimitsHysteresis#9 alarmHH');
    AssertEquals_BOOL(Expected := TRUE,
                      Actual := fbHighLimitsHysteresis.warnH,
                      Message := 'HighLimitsHysteresis#9 warnH');
    AssertEquals_BOOL(Expected := FALSE,
                      Actual := fbHighLimitsHysteresis.warnL,
                      Message := 'HighLimitsHysteresis#9 warnL');
    AssertEquals_BOOL(Expected := FALSE,
                      Actual := fbHighLimitsHysteresis.alarmLL,
                      Message := 'HighLimitsHysteresis#9 alarmLL');
    AssertEquals_WORD(Expected := 16#0021,
                      Actual := fbHighLimitsHysteresis.statusWord,
                      Message := 'HighLimitsHysteresis#9 statusWord');

    // #10, t = 900 мс — 11.0: H сброшен
    GVL_S7Clock.tSimNow := T#900MS;
    fbHighLimitsHysteresis.raw := 19008;
    fbHighLimitsHysteresis();
    AssertEquals_REAL(Expected := 11.0,
                      Actual := fbHighLimitsHysteresis.value,
                      Delta := 0.001,
                      Message := 'HighLimitsHysteresis#10 value');
    AssertEquals_BOOL(Expected := TRUE,
                      Actual := fbHighLimitsHysteresis.valid,
                      Message := 'HighLimitsHysteresis#10 valid');
    AssertEquals_BOOL(Expected := FALSE,
                      Actual := fbHighLimitsHysteresis.channelFault,
                      Message := 'HighLimitsHysteresis#10 channelFault');
    AssertEquals_BOOL(Expected := FALSE,
                      Actual := fbHighLimitsHysteresis.overrange,
                      Message := 'HighLimitsHysteresis#10 overrange');
    AssertEquals_BOOL(Expected := FALSE,
                      Actual := fbHighLimitsHysteresis.underrange,
                      Message := 'HighLimitsHysteresis#10 underrange');
    AssertEquals_BOOL(Expected := FALSE,
                      Actual := fbHighLimitsHysteresis.alarmHH,
                      Message := 'HighLimitsHysteresis#10 alarmHH');
    AssertEquals_BOOL(Expected := FALSE,
                      Actual := fbHighLimitsHysteresis.warnH,
                      Message := 'HighLimitsHysteresis#10 warnH');
    AssertEquals_BOOL(Expected := FALSE,
                      Actual := fbHighLimitsHysteresis.warnL,
                      Message := 'HighLimitsHysteresis#10 warnL');
    AssertEquals_BOOL(Expected := FALSE,
                      Actual := fbHighLimitsHysteresis.alarmLL,
                      Message := 'HighLimitsHysteresis#10 alarmLL');
    AssertEquals_WORD(Expected := 16#0001,
                      Actual := fbHighLimitsHysteresis.statusWord,
                      Message := 'HighLimitsHysteresis#10 statusWord');

    GVL_S7Clock.xSimulation := FALSE;
END_IF
coUnit.TEST_FINISHED();

(* ---- LowLimitsHysteresis.method.impl.st ---- *)
// AUTO-GENERATED — не редактировать: scenarios/FB_AnalogIn.csv, сценарий LowLimitsHysteresis
coUnit.TEST('LowLimitsHysteresis');
IF NOT xLowLimitsHysteresisDone THEN
    xLowLimitsHysteresisDone := TRUE;
    GVL_S7Clock.xSimulation := TRUE;

    // #1, t = 0 мс — 3.0 — выше нижних уставок
    GVL_S7Clock.tSimNow := T#0MS;
    fbLowLimitsHysteresis.raw := 5184;
    fbLowLimitsHysteresis.rangeLow := 0.0;
    fbLowLimitsHysteresis.rangeHigh := 16.0;
    fbLowLimitsHysteresis.limitHH := 14.0;
    fbLowLimitsHysteresis.limitH := 12.0;
    fbLowLimitsHysteresis.limitL := 2.0;
    fbLowLimitsHysteresis.limitLL := 1.0;
    fbLowLimitsHysteresis.hysteresis := 0.5;
    fbLowLimitsHysteresis.substitute := 0.0;
    fbLowLimitsHysteresis.simulation := FALSE;
    fbLowLimitsHysteresis.simValue := 0.0;
    fbLowLimitsHysteresis();
    AssertEquals_REAL(Expected := 3.0,
                      Actual := fbLowLimitsHysteresis.value,
                      Delta := 0.001,
                      Message := 'LowLimitsHysteresis#1 value');
    AssertEquals_BOOL(Expected := TRUE,
                      Actual := fbLowLimitsHysteresis.valid,
                      Message := 'LowLimitsHysteresis#1 valid');
    AssertEquals_BOOL(Expected := FALSE,
                      Actual := fbLowLimitsHysteresis.channelFault,
                      Message := 'LowLimitsHysteresis#1 channelFault');
    AssertEquals_BOOL(Expected := FALSE,
                      Actual := fbLowLimitsHysteresis.overrange,
                      Message := 'LowLimitsHysteresis#1 overrange');
    AssertEquals_BOOL(Expected := FALSE,
                      Actual := fbLowLimitsHysteresis.underrange,
                      Message := 'LowLimitsHysteresis#1 underrange');
    AssertEquals_BOOL(Expected := FALSE,
                      Actual := fbLowLimitsHysteresis.alarmHH,
                      Message := 'LowLimitsHysteresis#1 alarmHH');
    AssertEquals_BOOL(Expected := FALSE,
                      Actual := fbLowLimitsHysteresis.warnH,
                      Message := 'LowLimitsHysteresis#1 warnH');
    AssertEquals_BOOL(Expected := FALSE,
                      Actual := fbLowLimitsHysteresis.warnL,
                      Message := 'LowLimitsHysteresis#1 warnL');
    AssertEquals_BOOL(Expected := FALSE,
                      Actual := fbLowLimitsHysteresis.alarmLL,
                      Message := 'LowLimitsHysteresis#1 alarmLL');
    AssertEquals_WORD(Expected := 16#0001,
                      Actual := fbLowLimitsHysteresis.statusWord,
                      Message := 'LowLimitsHysteresis#1 statusWord');

    // #2, t = 100 мс — 2.0 = limitL: L включается
    GVL_S7Clock.tSimNow := T#100MS;
    fbLowLimitsHysteresis.raw := 3456;
    fbLowLimitsHysteresis();
    AssertEquals_REAL(Expected := 2.0,
                      Actual := fbLowLimitsHysteresis.value,
                      Delta := 0.001,
                      Message := 'LowLimitsHysteresis#2 value');
    AssertEquals_BOOL(Expected := TRUE,
                      Actual := fbLowLimitsHysteresis.valid,
                      Message := 'LowLimitsHysteresis#2 valid');
    AssertEquals_BOOL(Expected := FALSE,
                      Actual := fbLowLimitsHysteresis.channelFault,
                      Message := 'LowLimitsHysteresis#2 channelFault');
    AssertEquals_BOOL(Expected := FALSE,
                      Actual := fbLowLimitsHysteresis.overrange,
                      Message := 'LowLimitsHysteresis#2 overrange');
    AssertEquals_BOOL(Expected := FALSE,
                      Actual := fbLowLimitsHysteresis.underrange,
                      Message := 'LowLimitsHysteresis#2 underrange');
    AssertEquals_BOOL(Expected := FALSE,
                      Actual := fbLowLimitsHysteresis.alarmHH,
                      Message := 'LowLimitsHysteresis#2 alarmHH');
    AssertEquals_BOOL(Expected := FALSE,
                      Actual := fbLowLimitsHysteresis.warnH,
                      Message := 'LowLimitsHysteresis#2 warnH');
    AssertEquals_BOOL(Expected := TRUE,
                      Actual := fbLowLimitsHysteresis.warnL,
                      Message := 'LowLimitsHysteresis#2 warnL');
    AssertEquals_BOOL(Expected := FALSE,
                      Actual := fbLowLimitsHysteresis.alarmLL,
                      Message := 'LowLimitsHysteresis#2 alarmLL');
    AssertEquals_WORD(Expected := 16#0041,
                      Actual := fbLowLimitsHysteresis.statusWord,
                      Message := 'LowLimitsHysteresis#2 statusWord');

    // #3, t = 200 мс — 2.25 — в зоне гистерезиса, L держится
    GVL_S7Clock.tSimNow := T#200MS;
    fbLowLimitsHysteresis.raw := 3888;
    fbLowLimitsHysteresis();
    AssertEquals_REAL(Expected := 2.25,
                      Actual := fbLowLimitsHysteresis.value,
                      Delta := 0.001,
                      Message := 'LowLimitsHysteresis#3 value');
    AssertEquals_BOOL(Expected := TRUE,
                      Actual := fbLowLimitsHysteresis.valid,
                      Message := 'LowLimitsHysteresis#3 valid');
    AssertEquals_BOOL(Expected := FALSE,
                      Actual := fbLowLimitsHysteresis.channelFault,
                      Message := 'LowLimitsHysteresis#3 channelFault');
    AssertEquals_BOOL(Expected := FALSE,
                      Actual := fbLowLimitsHysteresis.overrange,
                      Message := 'LowLimitsHysteresis#3 overrange');
    AssertEquals_BOOL(Expected := FALSE,
                      Actual := fbLowLimitsHysteresis.underrange,
                      Message := 'LowLimitsHysteresis#3 underrange');
    AssertEquals_BOOL(Expected := FALSE,
                      Actual := fbLowLimitsHysteresis.alarmHH,
                      Message := 'LowLimitsHysteresis#3 alarmHH');
    AssertEquals_BOOL(Expected := FALSE,
                      Actual := fbLowLimitsHysteresis.warnH,
                      Message := 'LowLimitsHysteresis#3 warnH');
    AssertEquals_BOOL(Expected := TRUE,
                      Actual := fbLowLimitsHysteresis.warnL,
                      Message := 'LowLimitsHysteresis#3 warnL');
    AssertEquals_BOOL(Expected := FALSE,
                      Actual := fbLowLimitsHysteresis.alarmLL,
                      Message := 'LowLimitsHysteresis#3 alarmLL');
    AssertEquals_WORD(Expected := 16#0041,
                      Actual := fbLowLimitsHysteresis.statusWord,
                      Message := 'LowLimitsHysteresis#3 statusWord');

    // #4, t = 300 мс — 2.5 = limitL + hysteresis: не больше порога, L держится
    GVL_S7Clock.tSimNow := T#300MS;
    fbLowLimitsHysteresis.raw := 4320;
    fbLowLimitsHysteresis();
    AssertEquals_REAL(Expected := 2.5,
                      Actual := fbLowLimitsHysteresis.value,
                      Delta := 0.001,
                      Message := 'LowLimitsHysteresis#4 value');
    AssertEquals_BOOL(Expected := TRUE,
                      Actual := fbLowLimitsHysteresis.valid,
                      Message := 'LowLimitsHysteresis#4 valid');
    AssertEquals_BOOL(Expected := FALSE,
                      Actual := fbLowLimitsHysteresis.channelFault,
                      Message := 'LowLimitsHysteresis#4 channelFault');
    AssertEquals_BOOL(Expected := FALSE,
                      Actual := fbLowLimitsHysteresis.overrange,
                      Message := 'LowLimitsHysteresis#4 overrange');
    AssertEquals_BOOL(Expected := FALSE,
                      Actual := fbLowLimitsHysteresis.underrange,
                      Message := 'LowLimitsHysteresis#4 underrange');
    AssertEquals_BOOL(Expected := FALSE,
                      Actual := fbLowLimitsHysteresis.alarmHH,
                      Message := 'LowLimitsHysteresis#4 alarmHH');
    AssertEquals_BOOL(Expected := FALSE,
                      Actual := fbLowLimitsHysteresis.warnH,
                      Message := 'LowLimitsHysteresis#4 warnH');
    AssertEquals_BOOL(Expected := TRUE,
                      Actual := fbLowLimitsHysteresis.warnL,
                      Message := 'LowLimitsHysteresis#4 warnL');
    AssertEquals_BOOL(Expected := FALSE,
                      Actual := fbLowLimitsHysteresis.alarmLL,
                      Message := 'LowLimitsHysteresis#4 alarmLL');
    AssertEquals_WORD(Expected := 16#0041,
                      Actual := fbLowLimitsHysteresis.statusWord,
                      Message := 'LowLimitsHysteresis#4 statusWord');

    // #5, t = 400 мс — 2.75 > 2.5: L сбрасывается
    GVL_S7Clock.tSimNow := T#400MS;
    fbLowLimitsHysteresis.raw := 4752;
    fbLowLimitsHysteresis();
    AssertEquals_REAL(Expected := 2.75,
                      Actual := fbLowLimitsHysteresis.value,
                      Delta := 0.001,
                      Message := 'LowLimitsHysteresis#5 value');
    AssertEquals_BOOL(Expected := TRUE,
                      Actual := fbLowLimitsHysteresis.valid,
                      Message := 'LowLimitsHysteresis#5 valid');
    AssertEquals_BOOL(Expected := FALSE,
                      Actual := fbLowLimitsHysteresis.channelFault,
                      Message := 'LowLimitsHysteresis#5 channelFault');
    AssertEquals_BOOL(Expected := FALSE,
                      Actual := fbLowLimitsHysteresis.overrange,
                      Message := 'LowLimitsHysteresis#5 overrange');
    AssertEquals_BOOL(Expected := FALSE,
                      Actual := fbLowLimitsHysteresis.underrange,
                      Message := 'LowLimitsHysteresis#5 underrange');
    AssertEquals_BOOL(Expected := FALSE,
                      Actual := fbLowLimitsHysteresis.alarmHH,
                      Message := 'LowLimitsHysteresis#5 alarmHH');
    AssertEquals_BOOL(Expected := FALSE,
                      Actual := fbLowLimitsHysteresis.warnH,
                      Message := 'LowLimitsHysteresis#5 warnH');
    AssertEquals_BOOL(Expected := FALSE,
                      Actual := fbLowLimitsHysteresis.warnL,
                      Message := 'LowLimitsHysteresis#5 warnL');
    AssertEquals_BOOL(Expected := FALSE,
                      Actual := fbLowLimitsHysteresis.alarmLL,
                      Message := 'LowLimitsHysteresis#5 alarmLL');
    AssertEquals_WORD(Expected := 16#0001,
                      Actual := fbLowLimitsHysteresis.statusWord,
                      Message := 'LowLimitsHysteresis#5 statusWord');

    // #6, t = 500 мс — 1.0 = limitLL: L и LL
    GVL_S7Clock.tSimNow := T#500MS;
    fbLowLimitsHysteresis.raw := 1728;
    fbLowLimitsHysteresis();
    AssertEquals_REAL(Expected := 1.0,
                      Actual := fbLowLimitsHysteresis.value,
                      Delta := 0.001,
                      Message := 'LowLimitsHysteresis#6 value');
    AssertEquals_BOOL(Expected := TRUE,
                      Actual := fbLowLimitsHysteresis.valid,
                      Message := 'LowLimitsHysteresis#6 valid');
    AssertEquals_BOOL(Expected := FALSE,
                      Actual := fbLowLimitsHysteresis.channelFault,
                      Message := 'LowLimitsHysteresis#6 channelFault');
    AssertEquals_BOOL(Expected := FALSE,
                      Actual := fbLowLimitsHysteresis.overrange,
                      Message := 'LowLimitsHysteresis#6 overrange');
    AssertEquals_BOOL(Expected := FALSE,
                      Actual := fbLowLimitsHysteresis.underrange,
                      Message := 'LowLimitsHysteresis#6 underrange');
    AssertEquals_BOOL(Expected := FALSE,
                      Actual := fbLowLimitsHysteresis.alarmHH,
                      Message := 'LowLimitsHysteresis#6 alarmHH');
    AssertEquals_BOOL(Expected := FALSE,
                      Actual := fbLowLimitsHysteresis.warnH,
                      Message := 'LowLimitsHysteresis#6 warnH');
    AssertEquals_BOOL(Expected := TRUE,
                      Actual := fbLowLimitsHysteresis.warnL,
                      Message := 'LowLimitsHysteresis#6 warnL');
    AssertEquals_BOOL(Expected := TRUE,
                      Actual := fbLowLimitsHysteresis.alarmLL,
                      Message := 'LowLimitsHysteresis#6 alarmLL');
    AssertEquals_WORD(Expected := 16#00C1,
                      Actual := fbLowLimitsHysteresis.statusWord,
                      Message := 'LowLimitsHysteresis#6 statusWord');

    // #7, t = 600 мс — 1.5 = limitLL + hysteresis: LL держится
    GVL_S7Clock.tSimNow := T#600MS;
    fbLowLimitsHysteresis.raw := 2592;
    fbLowLimitsHysteresis();
    AssertEquals_REAL(Expected := 1.5,
                      Actual := fbLowLimitsHysteresis.value,
                      Delta := 0.001,
                      Message := 'LowLimitsHysteresis#7 value');
    AssertEquals_BOOL(Expected := TRUE,
                      Actual := fbLowLimitsHysteresis.valid,
                      Message := 'LowLimitsHysteresis#7 valid');
    AssertEquals_BOOL(Expected := FALSE,
                      Actual := fbLowLimitsHysteresis.channelFault,
                      Message := 'LowLimitsHysteresis#7 channelFault');
    AssertEquals_BOOL(Expected := FALSE,
                      Actual := fbLowLimitsHysteresis.overrange,
                      Message := 'LowLimitsHysteresis#7 overrange');
    AssertEquals_BOOL(Expected := FALSE,
                      Actual := fbLowLimitsHysteresis.underrange,
                      Message := 'LowLimitsHysteresis#7 underrange');
    AssertEquals_BOOL(Expected := FALSE,
                      Actual := fbLowLimitsHysteresis.alarmHH,
                      Message := 'LowLimitsHysteresis#7 alarmHH');
    AssertEquals_BOOL(Expected := FALSE,
                      Actual := fbLowLimitsHysteresis.warnH,
                      Message := 'LowLimitsHysteresis#7 warnH');
    AssertEquals_BOOL(Expected := TRUE,
                      Actual := fbLowLimitsHysteresis.warnL,
                      Message := 'LowLimitsHysteresis#7 warnL');
    AssertEquals_BOOL(Expected := TRUE,
                      Actual := fbLowLimitsHysteresis.alarmLL,
                      Message := 'LowLimitsHysteresis#7 alarmLL');
    AssertEquals_WORD(Expected := 16#00C1,
                      Actual := fbLowLimitsHysteresis.statusWord,
                      Message := 'LowLimitsHysteresis#7 statusWord');

    // #8, t = 700 мс — 1.75 > 1.5: LL сброшен; 1.75 <= 2.0 — L
    GVL_S7Clock.tSimNow := T#700MS;
    fbLowLimitsHysteresis.raw := 3024;
    fbLowLimitsHysteresis();
    AssertEquals_REAL(Expected := 1.75,
                      Actual := fbLowLimitsHysteresis.value,
                      Delta := 0.001,
                      Message := 'LowLimitsHysteresis#8 value');
    AssertEquals_BOOL(Expected := TRUE,
                      Actual := fbLowLimitsHysteresis.valid,
                      Message := 'LowLimitsHysteresis#8 valid');
    AssertEquals_BOOL(Expected := FALSE,
                      Actual := fbLowLimitsHysteresis.channelFault,
                      Message := 'LowLimitsHysteresis#8 channelFault');
    AssertEquals_BOOL(Expected := FALSE,
                      Actual := fbLowLimitsHysteresis.overrange,
                      Message := 'LowLimitsHysteresis#8 overrange');
    AssertEquals_BOOL(Expected := FALSE,
                      Actual := fbLowLimitsHysteresis.underrange,
                      Message := 'LowLimitsHysteresis#8 underrange');
    AssertEquals_BOOL(Expected := FALSE,
                      Actual := fbLowLimitsHysteresis.alarmHH,
                      Message := 'LowLimitsHysteresis#8 alarmHH');
    AssertEquals_BOOL(Expected := FALSE,
                      Actual := fbLowLimitsHysteresis.warnH,
                      Message := 'LowLimitsHysteresis#8 warnH');
    AssertEquals_BOOL(Expected := TRUE,
                      Actual := fbLowLimitsHysteresis.warnL,
                      Message := 'LowLimitsHysteresis#8 warnL');
    AssertEquals_BOOL(Expected := FALSE,
                      Actual := fbLowLimitsHysteresis.alarmLL,
                      Message := 'LowLimitsHysteresis#8 alarmLL');
    AssertEquals_WORD(Expected := 16#0041,
                      Actual := fbLowLimitsHysteresis.statusWord,
                      Message := 'LowLimitsHysteresis#8 statusWord');

    // #9, t = 800 мс — 1.25 > limitLL: LL не включается
    GVL_S7Clock.tSimNow := T#800MS;
    fbLowLimitsHysteresis.raw := 2160;
    fbLowLimitsHysteresis();
    AssertEquals_REAL(Expected := 1.25,
                      Actual := fbLowLimitsHysteresis.value,
                      Delta := 0.001,
                      Message := 'LowLimitsHysteresis#9 value');
    AssertEquals_BOOL(Expected := TRUE,
                      Actual := fbLowLimitsHysteresis.valid,
                      Message := 'LowLimitsHysteresis#9 valid');
    AssertEquals_BOOL(Expected := FALSE,
                      Actual := fbLowLimitsHysteresis.channelFault,
                      Message := 'LowLimitsHysteresis#9 channelFault');
    AssertEquals_BOOL(Expected := FALSE,
                      Actual := fbLowLimitsHysteresis.overrange,
                      Message := 'LowLimitsHysteresis#9 overrange');
    AssertEquals_BOOL(Expected := FALSE,
                      Actual := fbLowLimitsHysteresis.underrange,
                      Message := 'LowLimitsHysteresis#9 underrange');
    AssertEquals_BOOL(Expected := FALSE,
                      Actual := fbLowLimitsHysteresis.alarmHH,
                      Message := 'LowLimitsHysteresis#9 alarmHH');
    AssertEquals_BOOL(Expected := FALSE,
                      Actual := fbLowLimitsHysteresis.warnH,
                      Message := 'LowLimitsHysteresis#9 warnH');
    AssertEquals_BOOL(Expected := TRUE,
                      Actual := fbLowLimitsHysteresis.warnL,
                      Message := 'LowLimitsHysteresis#9 warnL');
    AssertEquals_BOOL(Expected := FALSE,
                      Actual := fbLowLimitsHysteresis.alarmLL,
                      Message := 'LowLimitsHysteresis#9 alarmLL');
    AssertEquals_WORD(Expected := 16#0041,
                      Actual := fbLowLimitsHysteresis.statusWord,
                      Message := 'LowLimitsHysteresis#9 statusWord');

    GVL_S7Clock.xSimulation := FALSE;
END_IF
coUnit.TEST_FINISHED();

(* ---- ScalingPoints.method.impl.st ---- *)
// AUTO-GENERATED — не редактировать: scenarios/FB_AnalogIn.csv, сценарий ScalingPoints
coUnit.TEST('ScalingPoints');
IF NOT xScalingPointsDone THEN
    xScalingPointsDone := TRUE;
    GVL_S7Clock.xSimulation := TRUE;

    // #1, t = 0 мс — 0 -> 0.0 бар; ниже L и LL
    GVL_S7Clock.tSimNow := T#0MS;
    fbScalingPoints.raw := 0;
    fbScalingPoints.rangeLow := 0.0;
    fbScalingPoints.rangeHigh := 16.0;
    fbScalingPoints.limitHH := 14.0;
    fbScalingPoints.limitH := 12.0;
    fbScalingPoints.limitL := 2.0;
    fbScalingPoints.limitLL := 1.0;
    fbScalingPoints.hysteresis := 0.5;
    fbScalingPoints.substitute := 0.0;
    fbScalingPoints.simulation := FALSE;
    fbScalingPoints.simValue := 0.0;
    fbScalingPoints();
    AssertEquals_REAL(Expected := 0.0,
                      Actual := fbScalingPoints.value,
                      Delta := 0.001,
                      Message := 'ScalingPoints#1 value');
    AssertEquals_BOOL(Expected := TRUE, Actual := fbScalingPoints.valid, Message := 'ScalingPoints#1 valid');
    AssertEquals_BOOL(Expected := FALSE,
                      Actual := fbScalingPoints.channelFault,
                      Message := 'ScalingPoints#1 channelFault');
    AssertEquals_BOOL(Expected := FALSE, Actual := fbScalingPoints.overrange, Message := 'ScalingPoints#1 overrange');
    AssertEquals_BOOL(Expected := FALSE, Actual := fbScalingPoints.underrange, Message := 'ScalingPoints#1 underrange');
    AssertEquals_BOOL(Expected := FALSE, Actual := fbScalingPoints.alarmHH, Message := 'ScalingPoints#1 alarmHH');
    AssertEquals_BOOL(Expected := FALSE, Actual := fbScalingPoints.warnH, Message := 'ScalingPoints#1 warnH');
    AssertEquals_BOOL(Expected := TRUE, Actual := fbScalingPoints.warnL, Message := 'ScalingPoints#1 warnL');
    AssertEquals_BOOL(Expected := TRUE, Actual := fbScalingPoints.alarmLL, Message := 'ScalingPoints#1 alarmLL');
    AssertEquals_WORD(Expected := 16#00C1,
                      Actual := fbScalingPoints.statusWord,
                      Message := 'ScalingPoints#1 statusWord');

    // #2, t = 100 мс — середина шкалы -> 8.0; L и LL сброшены (8.0 > 2.5 и > 1.5)
    GVL_S7Clock.tSimNow := T#100MS;
    fbScalingPoints.raw := 13824;
    fbScalingPoints();
    AssertEquals_REAL(Expected := 8.0,
                      Actual := fbScalingPoints.value,
                      Delta := 0.001,
                      Message := 'ScalingPoints#2 value');
    AssertEquals_BOOL(Expected := TRUE, Actual := fbScalingPoints.valid, Message := 'ScalingPoints#2 valid');
    AssertEquals_BOOL(Expected := FALSE,
                      Actual := fbScalingPoints.channelFault,
                      Message := 'ScalingPoints#2 channelFault');
    AssertEquals_BOOL(Expected := FALSE, Actual := fbScalingPoints.overrange, Message := 'ScalingPoints#2 overrange');
    AssertEquals_BOOL(Expected := FALSE, Actual := fbScalingPoints.underrange, Message := 'ScalingPoints#2 underrange');
    AssertEquals_BOOL(Expected := FALSE, Actual := fbScalingPoints.alarmHH, Message := 'ScalingPoints#2 alarmHH');
    AssertEquals_BOOL(Expected := FALSE, Actual := fbScalingPoints.warnH, Message := 'ScalingPoints#2 warnH');
    AssertEquals_BOOL(Expected := FALSE, Actual := fbScalingPoints.warnL, Message := 'ScalingPoints#2 warnL');
    AssertEquals_BOOL(Expected := FALSE, Actual := fbScalingPoints.alarmLL, Message := 'ScalingPoints#2 alarmLL');
    AssertEquals_WORD(Expected := 16#0001,
                      Actual := fbScalingPoints.statusWord,
                      Message := 'ScalingPoints#2 statusWord');

    // #3, t = 200 мс — номинальный максимум -> 16.0; HH и H
    GVL_S7Clock.tSimNow := T#200MS;
    fbScalingPoints.raw := 27648;
    fbScalingPoints();
    AssertEquals_REAL(Expected := 16.0,
                      Actual := fbScalingPoints.value,
                      Delta := 0.001,
                      Message := 'ScalingPoints#3 value');
    AssertEquals_BOOL(Expected := TRUE, Actual := fbScalingPoints.valid, Message := 'ScalingPoints#3 valid');
    AssertEquals_BOOL(Expected := FALSE,
                      Actual := fbScalingPoints.channelFault,
                      Message := 'ScalingPoints#3 channelFault');
    AssertEquals_BOOL(Expected := FALSE, Actual := fbScalingPoints.overrange, Message := 'ScalingPoints#3 overrange');
    AssertEquals_BOOL(Expected := FALSE, Actual := fbScalingPoints.underrange, Message := 'ScalingPoints#3 underrange');
    AssertEquals_BOOL(Expected := TRUE, Actual := fbScalingPoints.alarmHH, Message := 'ScalingPoints#3 alarmHH');
    AssertEquals_BOOL(Expected := TRUE, Actual := fbScalingPoints.warnH, Message := 'ScalingPoints#3 warnH');
    AssertEquals_BOOL(Expected := FALSE, Actual := fbScalingPoints.warnL, Message := 'ScalingPoints#3 warnL');
    AssertEquals_BOOL(Expected := FALSE, Actual := fbScalingPoints.alarmLL, Message := 'ScalingPoints#3 alarmLL');
    AssertEquals_WORD(Expected := 16#0031,
                      Actual := fbScalingPoints.statusWord,
                      Message := 'ScalingPoints#3 statusWord');

    // #4, t = 300 мс — четверть -> 4.0; HH и H сброшены
    GVL_S7Clock.tSimNow := T#300MS;
    fbScalingPoints.raw := 6912;
    fbScalingPoints();
    AssertEquals_REAL(Expected := 4.0,
                      Actual := fbScalingPoints.value,
                      Delta := 0.001,
                      Message := 'ScalingPoints#4 value');
    AssertEquals_BOOL(Expected := TRUE, Actual := fbScalingPoints.valid, Message := 'ScalingPoints#4 valid');
    AssertEquals_BOOL(Expected := FALSE,
                      Actual := fbScalingPoints.channelFault,
                      Message := 'ScalingPoints#4 channelFault');
    AssertEquals_BOOL(Expected := FALSE, Actual := fbScalingPoints.overrange, Message := 'ScalingPoints#4 overrange');
    AssertEquals_BOOL(Expected := FALSE, Actual := fbScalingPoints.underrange, Message := 'ScalingPoints#4 underrange');
    AssertEquals_BOOL(Expected := FALSE, Actual := fbScalingPoints.alarmHH, Message := 'ScalingPoints#4 alarmHH');
    AssertEquals_BOOL(Expected := FALSE, Actual := fbScalingPoints.warnH, Message := 'ScalingPoints#4 warnH');
    AssertEquals_BOOL(Expected := FALSE, Actual := fbScalingPoints.warnL, Message := 'ScalingPoints#4 warnL');
    AssertEquals_BOOL(Expected := FALSE, Actual := fbScalingPoints.alarmLL, Message := 'ScalingPoints#4 alarmLL');
    AssertEquals_WORD(Expected := 16#0001,
                      Actual := fbScalingPoints.statusWord,
                      Message := 'ScalingPoints#4 statusWord');

    // #5, t = 400 мс — -> 12.0 = limitH: H включается (>=)
    GVL_S7Clock.tSimNow := T#400MS;
    fbScalingPoints.raw := 20736;
    fbScalingPoints();
    AssertEquals_REAL(Expected := 12.0,
                      Actual := fbScalingPoints.value,
                      Delta := 0.001,
                      Message := 'ScalingPoints#5 value');
    AssertEquals_BOOL(Expected := TRUE, Actual := fbScalingPoints.valid, Message := 'ScalingPoints#5 valid');
    AssertEquals_BOOL(Expected := FALSE,
                      Actual := fbScalingPoints.channelFault,
                      Message := 'ScalingPoints#5 channelFault');
    AssertEquals_BOOL(Expected := FALSE, Actual := fbScalingPoints.overrange, Message := 'ScalingPoints#5 overrange');
    AssertEquals_BOOL(Expected := FALSE, Actual := fbScalingPoints.underrange, Message := 'ScalingPoints#5 underrange');
    AssertEquals_BOOL(Expected := FALSE, Actual := fbScalingPoints.alarmHH, Message := 'ScalingPoints#5 alarmHH');
    AssertEquals_BOOL(Expected := TRUE, Actual := fbScalingPoints.warnH, Message := 'ScalingPoints#5 warnH');
    AssertEquals_BOOL(Expected := FALSE, Actual := fbScalingPoints.warnL, Message := 'ScalingPoints#5 warnL');
    AssertEquals_BOOL(Expected := FALSE, Actual := fbScalingPoints.alarmLL, Message := 'ScalingPoints#5 alarmLL');
    AssertEquals_WORD(Expected := 16#0021,
                      Actual := fbScalingPoints.statusWord,
                      Message := 'ScalingPoints#5 statusWord');

    // #6, t = 500 мс — -> 1.0 = limitLL: L и LL включаются (<=), H сброшен
    GVL_S7Clock.tSimNow := T#500MS;
    fbScalingPoints.raw := 1728;
    fbScalingPoints();
    AssertEquals_REAL(Expected := 1.0,
                      Actual := fbScalingPoints.value,
                      Delta := 0.001,
                      Message := 'ScalingPoints#6 value');
    AssertEquals_BOOL(Expected := TRUE, Actual := fbScalingPoints.valid, Message := 'ScalingPoints#6 valid');
    AssertEquals_BOOL(Expected := FALSE,
                      Actual := fbScalingPoints.channelFault,
                      Message := 'ScalingPoints#6 channelFault');
    AssertEquals_BOOL(Expected := FALSE, Actual := fbScalingPoints.overrange, Message := 'ScalingPoints#6 overrange');
    AssertEquals_BOOL(Expected := FALSE, Actual := fbScalingPoints.underrange, Message := 'ScalingPoints#6 underrange');
    AssertEquals_BOOL(Expected := FALSE, Actual := fbScalingPoints.alarmHH, Message := 'ScalingPoints#6 alarmHH');
    AssertEquals_BOOL(Expected := FALSE, Actual := fbScalingPoints.warnH, Message := 'ScalingPoints#6 warnH');
    AssertEquals_BOOL(Expected := TRUE, Actual := fbScalingPoints.warnL, Message := 'ScalingPoints#6 warnL');
    AssertEquals_BOOL(Expected := TRUE, Actual := fbScalingPoints.alarmLL, Message := 'ScalingPoints#6 alarmLL');
    AssertEquals_WORD(Expected := 16#00C1,
                      Actual := fbScalingPoints.statusWord,
                      Message := 'ScalingPoints#6 statusWord');

    GVL_S7Clock.xSimulation := FALSE;
END_IF
coUnit.TEST_FINISHED();

(* ---- Simulation.method.impl.st ---- *)
// AUTO-GENERATED — не редактировать: scenarios/FB_AnalogIn.csv, сценарий Simulation
coUnit.TEST('Simulation');
IF NOT xSimulationDone THEN
    xSimulationDone := TRUE;
    GVL_S7Clock.xSimulation := TRUE;

    // #1, t = 0 мс — неисправность, value = substitute 0.0
    GVL_S7Clock.tSimNow := T#0MS;
    fbSimulation.raw := 32767;
    fbSimulation.rangeLow := 0.0;
    fbSimulation.rangeHigh := 16.0;
    fbSimulation.limitHH := 14.0;
    fbSimulation.limitH := 12.0;
    fbSimulation.limitL := 2.0;
    fbSimulation.limitLL := 1.0;
    fbSimulation.hysteresis := 0.5;
    fbSimulation.substitute := 0.0;
    fbSimulation.simulation := FALSE;
    fbSimulation.simValue := 0.0;
    fbSimulation();
    AssertEquals_REAL(Expected := 0.0, Actual := fbSimulation.value, Delta := 0.001, Message := 'Simulation#1 value');
    AssertEquals_BOOL(Expected := FALSE, Actual := fbSimulation.valid, Message := 'Simulation#1 valid');
    AssertEquals_BOOL(Expected := TRUE, Actual := fbSimulation.channelFault, Message := 'Simulation#1 channelFault');
    AssertEquals_BOOL(Expected := FALSE, Actual := fbSimulation.overrange, Message := 'Simulation#1 overrange');
    AssertEquals_BOOL(Expected := FALSE, Actual := fbSimulation.underrange, Message := 'Simulation#1 underrange');
    AssertEquals_BOOL(Expected := FALSE, Actual := fbSimulation.alarmHH, Message := 'Simulation#1 alarmHH');
    AssertEquals_BOOL(Expected := FALSE, Actual := fbSimulation.warnH, Message := 'Simulation#1 warnH');
    AssertEquals_BOOL(Expected := FALSE, Actual := fbSimulation.warnL, Message := 'Simulation#1 warnL');
    AssertEquals_BOOL(Expected := FALSE, Actual := fbSimulation.alarmLL, Message := 'Simulation#1 alarmLL');
    AssertEquals_WORD(Expected := 16#0002, Actual := fbSimulation.statusWord, Message := 'Simulation#1 statusWord');

    // #2, t = 100 мс — имитация 15.0: valid, HH и H; channelFault по raw остаётся
    GVL_S7Clock.tSimNow := T#100MS;
    fbSimulation.simulation := TRUE;
    fbSimulation.simValue := 15.0;
    fbSimulation();
    AssertEquals_REAL(Expected := 15.0, Actual := fbSimulation.value, Delta := 0.001, Message := 'Simulation#2 value');
    AssertEquals_BOOL(Expected := TRUE, Actual := fbSimulation.valid, Message := 'Simulation#2 valid');
    AssertEquals_BOOL(Expected := TRUE, Actual := fbSimulation.channelFault, Message := 'Simulation#2 channelFault');
    AssertEquals_BOOL(Expected := FALSE, Actual := fbSimulation.overrange, Message := 'Simulation#2 overrange');
    AssertEquals_BOOL(Expected := FALSE, Actual := fbSimulation.underrange, Message := 'Simulation#2 underrange');
    AssertEquals_BOOL(Expected := TRUE, Actual := fbSimulation.alarmHH, Message := 'Simulation#2 alarmHH');
    AssertEquals_BOOL(Expected := TRUE, Actual := fbSimulation.warnH, Message := 'Simulation#2 warnH');
    AssertEquals_BOOL(Expected := FALSE, Actual := fbSimulation.warnL, Message := 'Simulation#2 warnL');
    AssertEquals_BOOL(Expected := FALSE, Actual := fbSimulation.alarmLL, Message := 'Simulation#2 alarmLL');
    AssertEquals_WORD(Expected := 16#0133, Actual := fbSimulation.statusWord, Message := 'Simulation#2 statusWord');

    // #3, t = 200 мс — 13.0 < 13.5: HH сброшен, H держится
    GVL_S7Clock.tSimNow := T#200MS;
    fbSimulation.simValue := 13.0;
    fbSimulation();
    AssertEquals_REAL(Expected := 13.0, Actual := fbSimulation.value, Delta := 0.001, Message := 'Simulation#3 value');
    AssertEquals_BOOL(Expected := TRUE, Actual := fbSimulation.valid, Message := 'Simulation#3 valid');
    AssertEquals_BOOL(Expected := TRUE, Actual := fbSimulation.channelFault, Message := 'Simulation#3 channelFault');
    AssertEquals_BOOL(Expected := FALSE, Actual := fbSimulation.overrange, Message := 'Simulation#3 overrange');
    AssertEquals_BOOL(Expected := FALSE, Actual := fbSimulation.underrange, Message := 'Simulation#3 underrange');
    AssertEquals_BOOL(Expected := FALSE, Actual := fbSimulation.alarmHH, Message := 'Simulation#3 alarmHH');
    AssertEquals_BOOL(Expected := TRUE, Actual := fbSimulation.warnH, Message := 'Simulation#3 warnH');
    AssertEquals_BOOL(Expected := FALSE, Actual := fbSimulation.warnL, Message := 'Simulation#3 warnL');
    AssertEquals_BOOL(Expected := FALSE, Actual := fbSimulation.alarmLL, Message := 'Simulation#3 alarmLL');
    AssertEquals_WORD(Expected := 16#0123, Actual := fbSimulation.statusWord, Message := 'Simulation#3 statusWord');

    // #4, t = 300 мс — канал исправен, имитация продолжается: value 13.0
    GVL_S7Clock.tSimNow := T#300MS;
    fbSimulation.raw := 13824;
    fbSimulation();
    AssertEquals_REAL(Expected := 13.0, Actual := fbSimulation.value, Delta := 0.001, Message := 'Simulation#4 value');
    AssertEquals_BOOL(Expected := TRUE, Actual := fbSimulation.valid, Message := 'Simulation#4 valid');
    AssertEquals_BOOL(Expected := FALSE, Actual := fbSimulation.channelFault, Message := 'Simulation#4 channelFault');
    AssertEquals_BOOL(Expected := FALSE, Actual := fbSimulation.overrange, Message := 'Simulation#4 overrange');
    AssertEquals_BOOL(Expected := FALSE, Actual := fbSimulation.underrange, Message := 'Simulation#4 underrange');
    AssertEquals_BOOL(Expected := FALSE, Actual := fbSimulation.alarmHH, Message := 'Simulation#4 alarmHH');
    AssertEquals_BOOL(Expected := TRUE, Actual := fbSimulation.warnH, Message := 'Simulation#4 warnH');
    AssertEquals_BOOL(Expected := FALSE, Actual := fbSimulation.warnL, Message := 'Simulation#4 warnL');
    AssertEquals_BOOL(Expected := FALSE, Actual := fbSimulation.alarmLL, Message := 'Simulation#4 alarmLL');
    AssertEquals_WORD(Expected := 16#0121, Actual := fbSimulation.statusWord, Message := 'Simulation#4 statusWord');

    // #5, t = 400 мс — имитация снята: value по raw 8.0, H сброшен
    GVL_S7Clock.tSimNow := T#400MS;
    fbSimulation.simulation := FALSE;
    fbSimulation();
    AssertEquals_REAL(Expected := 8.0, Actual := fbSimulation.value, Delta := 0.001, Message := 'Simulation#5 value');
    AssertEquals_BOOL(Expected := TRUE, Actual := fbSimulation.valid, Message := 'Simulation#5 valid');
    AssertEquals_BOOL(Expected := FALSE, Actual := fbSimulation.channelFault, Message := 'Simulation#5 channelFault');
    AssertEquals_BOOL(Expected := FALSE, Actual := fbSimulation.overrange, Message := 'Simulation#5 overrange');
    AssertEquals_BOOL(Expected := FALSE, Actual := fbSimulation.underrange, Message := 'Simulation#5 underrange');
    AssertEquals_BOOL(Expected := FALSE, Actual := fbSimulation.alarmHH, Message := 'Simulation#5 alarmHH');
    AssertEquals_BOOL(Expected := FALSE, Actual := fbSimulation.warnH, Message := 'Simulation#5 warnH');
    AssertEquals_BOOL(Expected := FALSE, Actual := fbSimulation.warnL, Message := 'Simulation#5 warnL');
    AssertEquals_BOOL(Expected := FALSE, Actual := fbSimulation.alarmLL, Message := 'Simulation#5 alarmLL');
    AssertEquals_WORD(Expected := 16#0001, Actual := fbSimulation.statusWord, Message := 'Simulation#5 statusWord');

    GVL_S7Clock.xSimulation := FALSE;
END_IF
coUnit.TEST_FINISHED();
